Fanuc KAREL source: kt00332.KL

-- PROVISIONAL review KL for V940-1; original PC SHA256 b3069f6366886043a367c5c37da46066d7e6a751381f3a15e8b1443fb4cba0a9
-- Incomplete behavior may be omitted. Consult companion uncertainty JSON. Do not deploy.
PROGRAM KT00332
%NOLOCKGROUP
VAR
  I1 : INTEGER
  OUT : BOOLEAN
-- UNRESOLVED_DECL H2 type=002017
BEGIN
  -- V9_ZERO_TABLE_METADATA_HINT layout=0001; no indexed target words; source/name/runtime held
  -- UNRESOLVED_PC offsets 5-16; opcodes 2E,23
  -- UNRESOLVED_PC offsets 21-35; opcodes 2E,22,9D,33,B4
  -- UNRESOLVED_PC offsets 40-62; opcodes 21,22,9D,33,B3,59,23
  -- UNRESOLVED_PC offsets 67-71; opcodes 7F
END KT00332
